FUNCTION F_BuildAPTitle : STRING
VAR_INPUT
    iValue : UDINT;
END_VAR

F_BuildAPTitle := CONCAT('1.1.1.999.', UDINT_TO_STRING(iValue));

END_FUNCTION

(* stored: Version 1.1.0.1
   POU F_BuildAPTitle: Id {059a3f35-772f-419b-9c48-7518e55ff3d9}, SpecialFunc None *)
